TYPE "ST_UnitProbeStationCfg"
VERSION : 0.1
   STRUCT
      "SchemaVersion" : UInt := 2;
      "SiteLabel" : String[80] := 'bench';
      "Enabled" : Bool := TRUE;
      "LongText" : String[80] := 'long default';
   END_STRUCT;
END_TYPE
